(* Simple 2-state coating selector, no PMPS: thin ND-framework wrapper
   around FB_PositionStateND, ported from a deprecated EXTENDS
   FB_PositionStateBase device. Single motor, no beam-safety gating.

   The integrator supplies sName/fPosition/fDelta/nEncoderCount for
   every state via FB_CC_StateDefaultsConfig (Convention B, the same
   split FB_SXR_SATT_Stage uses). This FB owns none of that config
   itself. FB_KBO_Coating_States uses the other split (Convention A,
   device owns sName/fDelta). Motor and state array are caller-owned,
   injected via FB_Init. *)
{attribute 'call_after_init'}
FUNCTION_BLOCK FB_Coating_States_NoPMPS
VAR
    (* State-enum bridge bound to FB_PositionStateND's REFERENCE TO UINT
       param via the shared UINT base. EPICS owns it through the pytmc
       pragma; PLC code must go through the EnumSet property instead of
       touching it directly. *)
    // Set this to a non-unknown value to request a new move.
    {attribute 'pytmc' := '
        pv: SET
        io: io
    '}
    eEnumSet : E_Coating_States;
    {attribute 'no_copy'}
    aiMotionStage    : REFERENCE TO ARRAY[1..MotionConstants.MAX_STATE_MOTORS] OF I_MotionStage;
    {attribute 'no_copy'}
    astPositionState : REFERENCE TO ARRAY[1..MotionConstants.MAX_STATE_MOTORS]
                                         OF ARRAY[1..GeneralConstants.MAX_STATES] OF ST_PositionState;

    bEnableMotion : BOOL := TRUE;

    {attribute 'pytmc' := 'pv: MMS'}
    fbStates : FB_PositionStateND(
        aiMotionStage        := aiMotionStage,
        astPositionState     := astPositionState,
        nActiveMotorCount    := 1,
        eEnumSet             := eEnumSet,
        eEnumGet             := eEnumGet,
        bEnableMotion        := bEnableMotion,
        eMotionRequestPolicy := E_MotionRequestPolicy.INTERRUPT
    );
END_VAR
VAR_OUTPUT
    // The current position state as an enum.
    {attribute 'pytmc' := '
        pv: GET
        io: i
    '}
    eEnumGet : E_Coating_States;
END_VAR

IF NOT __ISVALIDREF(aiMotionStage)
   OR NOT __ISVALIDREF(astPositionState) THEN
    RETURN;
END_IF

fbStates();


{attribute 'call_after_init'}
METHOD CallAfterInit
THIS^.fbStates.CallAfterInitStateMover(
    aiMotionStage         := aiMotionStage,
    astPositionState      := astPositionState,
    nActiveMotorCount     := 1,
    eEnumSet              := eEnumSet,
    eEnumGet              := eEnumGet,
    bEnableMotion         := bEnableMotion,
    eMotionRequestPolicy  := E_MotionRequestPolicy.INTERRUPT,
);
END_METHOD


METHOD FB_Init: BOOL
VAR_INPUT
    bInitRetains: BOOL; // TRUE: the retain variables are initialized (reset warm / reset cold)
    bInCopyCode: BOOL;  // TRUE: the instance will be copied to the copy code afterward (online change)
    aiMotionStage    : REFERENCE TO ARRAY[1..MotionConstants.MAX_STATE_MOTORS] OF I_MotionStage;
    astPositionState : REFERENCE TO ARRAY[1..MotionConstants.MAX_STATE_MOTORS]
                                         OF ARRAY[1..GeneralConstants.MAX_STATES] OF ST_PositionState;
END_VAR
THIS^.aiMotionStage    REF= aiMotionStage;
THIS^.astPositionState REF= astPositionState;
END_METHOD

(* Current position state. Read-only; written by the state mover. *)
PROPERTY EnumGet : E_Coating_States
GET
EnumGet := eEnumGet;
END_GET
END_PROPERTY

(* Request a new move, e.g. `fbCoating.EnumSet := E_Coating_States.Coating2;`.
   The state mover consumes and clears the request. *)
PROPERTY EnumSet : E_Coating_States
GET
EnumSet := eEnumSet;
END_GET
SET
eEnumSet := EnumSet;
END_SET
END_PROPERTY

END_FUNCTION_BLOCK

(* stored: Version 1.1.0.1
   POU FB_Coating_States_NoPMPS: Id {5e9b2f4d-8c6a-4b1e-93d7-1f4a2c6e9b05}, SpecialFunc None
   Method CallAfterInit: Id {5e9b2f4d-8c6a-4b1e-93d7-1f4a2c6e9b06}
   Method FB_Init: Id {5e9b2f4d-8c6a-4b1e-93d7-1f4a2c6e9b07}
   Property EnumGet: Id {82900509-1fb4-4919-9e80-5962027d071a}
   Get Get: Id {39def1cf-6f28-4f13-9acb-27339259f10b}
   Property EnumSet: Id {9c11b2da-dab1-4f61-9973-46a58278635f}
   Get Get: Id {8e4b8823-1c26-481c-99b9-da1f4f4ee831}
   Set Set: Id {ee289a61-67ea-4545-8d3c-adce6c116fda} *)
